// TIA Portal V20 export
DATA_BLOCK "DB_STS_M"   // DB101
{ S7_Optimized_Access := 'FALSE' }
// stored: AutoNumber false
   VAR
      OP0 : Struct
         STS_M0 : UInt;
         STS_M1 : UInt;
         STS_M2 : UInt;
         STS_M3 : UInt;
         STS_M4 : UInt;
         STS_M5 : UInt;
         STS_M6 : UInt;
         STS_M7 : UInt;
         STS_M8 : UInt;
         STS_M9 : UInt;
         STS_M10 : UInt;
         STS_M11 : UInt;
         STS_M12 : UInt;
         STS_M13 : UInt;
         STS_M14 : UInt;
         STS_M15 : UInt;
      END_STRUCT;
      OP1 : Struct
         KARUSEL : UInt;
         ZARAZKA : UInt;
         STS_M2 : UInt;
         STS_M3 : UInt;
         STS_M4 : UInt;
         STS_M5 : UInt;
         STS_M6 : UInt;
         STS_M7 : UInt;
         STS_M8 : UInt;
         STS_M9 : UInt;
         STS_M10 : UInt;
         STS_M11 : UInt;
         STS_M12 : UInt;
         STS_M13 : UInt;
         STS_M14 : UInt;
         STS_M15 : UInt;
         OP1 : Struct
            STS_M0 : UInt;
            STS_M1 : UInt;
            STS_M2 : UInt;
            STS_M3 : UInt;
            STS_M4 : UInt;
            STS_M5 : UInt;
            STS_M6 : UInt;
            STS_M7 : UInt;
            STS_M8 : UInt;
            STS_M9 : UInt;
            STS_M10 : UInt;
            STS_M11 : UInt;
            STS_M12 : UInt;
            STS_M13 : UInt;
            STS_M14 : UInt;
            STS_M15 : UInt;
         END_STRUCT;
      END_STRUCT;
      OP2 : Struct
         A1 : UInt;
         A2 : UInt;
         A3 : UInt;
         A4 : UInt;
         A5 : UInt;
         A6 : UInt;
         A7 : UInt;
         A8 : UInt;
         STS_M8 : UInt;
         STS_M9 : UInt;
         STS_M10 : UInt;
         STS_M11 : UInt;
         STS_M12 : UInt;
         STS_M13 : UInt;
         STS_M14 : UInt;
         STS_M15 : UInt;
      END_STRUCT;
      OP3 : Struct
         B1 : UInt;
         B2 : UInt;
         B3 : UInt;
         B4 : UInt;
         B5 : UInt;
         B6 : UInt;
         B7 : UInt;
         B8 : UInt;
         STS_M8 : UInt;
         STS_M9 : UInt;
         STS_M10 : UInt;
         STS_M11 : UInt;
         STS_M12 : UInt;
         STS_M13 : UInt;
         STS_M14 : UInt;
         STS_M15 : UInt;
      END_STRUCT;
   END_VAR
BEGIN
END_DATA_BLOCK
